TYPE "DT_PAR_GEN_MEAS_2"
VERSION : 0.1
   STRUCT
      OIL_NDE_TEMP_VAL_LOW { S7_SetPoint := 'False'} : "DT_PARAM_SOLO" := (FALSE, 320, 0, 0.0, 0, T#0MS, 0.0, 0.0, '°C');
      OIL_NDE_TEMP_VAL_HIGH { S7_SetPoint := 'False'} : "DT_PARAM_SOLO" := (FALSE, 321, 0, 150.0, 0, T#0MS, 0.0, 0.0, '°C');
      OIL_NDE_TEMP_SCAL_FACTOR { S7_SetPoint := 'False'} : "DT_PARAM_SOLO" := (FALSE, 322, 0, 1.0, 0, T#0MS, 0.0, 0.0, '°C');
      OIL_NDE_TEMP_OFFSET { S7_SetPoint := 'False'} : "DT_PARAM_SOLO" := (FALSE, 323, 0, 0.0, 0, T#0MS, 0.0, 0.0, '°C');
      OIL_NDE_TEMP_H { S7_SetPoint := 'False'} : "DT_PARAM_SOLO" := (FALSE, 324, 0, 120.0, 0, T#0MS, 0.0, 0.0, '°C');
      OIL_NDE_TEMP_HH { S7_SetPoint := 'False'} : "DT_PARAM_SOLO" := (FALSE, 325, 0, 130.0, 0, T#0MS, 0.0, 0.0, '°C');
      THRUST_NDE_TEMP_VAL_LOW { S7_SetPoint := 'False'} : "DT_PARAM_SOLO" := (FALSE, 326, 0, 1.0, 0, T#0MS, 0.0, 0.0, '°C');
      THRUST_NDE_TEMP_VAL_HIGH { S7_SetPoint := 'False'} : "DT_PARAM_SOLO" := (FALSE, 327, 0, 0.0, 0, T#0MS, 0.0, 0.0, '°C');
      THRUST_NDE_TEMP_SCAL_FACTOR { S7_SetPoint := 'False'} : "DT_PARAM_SOLO" := (FALSE, 328, 0, 1.0, 0, T#0MS, 0.0, 0.0, '°C');
      THRUST_NDE_TEMP_OFFSET { S7_SetPoint := 'False'} : "DT_PARAM_SOLO" := (FALSE, 329, 0, 0.0, 0, T#0MS, 0.0, 0.0, '°C');
      THRUST_NDE_TEMP_H { S7_SetPoint := 'False'} : "DT_PARAM_SOLO" := (FALSE, 330, 0, 70.0, 0, T#0MS, 0.0, 0.0, '°C');
      THRUST_NDE_TEMP_HH { S7_SetPoint := 'False'} : "DT_PARAM_SOLO" := (FALSE, 331, 0, 80.0, 0, T#0MS, 0.0, 0.0, '°C');
      PARAM_12 { S7_SetPoint := 'False'} : "DT_PARAM_SOLO" := (FALSE, 332, 0, 0.0, 0, T#0MS, 0.0, 0.0, '');
      PARAM_13 { S7_SetPoint := 'False'} : "DT_PARAM_SOLO" := (FALSE, 333, 0, 120.0, 0, T#0MS, 0.0, 0.0, '');
      PARAM_14 { S7_SetPoint := 'False'} : "DT_PARAM_SOLO" := (FALSE, 334, 0, 1.0, 0, T#0MS, 0.0, 0.0, '');
      PARAM_15 { S7_SetPoint := 'False'} : "DT_PARAM_SOLO" := (FALSE, 335, 0, 0.0, 0, T#0MS, 0.0, 0.0, '');
      PARAM_16 { S7_SetPoint := 'False'} : "DT_PARAM_SOLO" := (FALSE, 336, 0, 70.0, 0, T#0MS, 0.0, 0.0, '');
      PARAM_17 { S7_SetPoint := 'False'} : "DT_PARAM_SOLO" := (FALSE, 337, 0, 80.0, 0, T#0MS, 0.0, 0.0, '');
      PARAM_18 { S7_SetPoint := 'False'} : "DT_PARAM_SOLO" := (FALSE, 338, 0, 0.0, 0, T#0MS, 0.0, 0.0, '');
      PARAM_19 { S7_SetPoint := 'False'} : "DT_PARAM_SOLO" := (FALSE, 339, 0, 0.0, 0, T#0MS, 0.0, 0.0, '');
      PARAM_20 { S7_SetPoint := 'False'} : "DT_PARAM_SOLO" := (FALSE, 340, 0, 0.0, 0, T#0MS, 0.0, 0.0, '');
      PARAM_21 { S7_SetPoint := 'False'} : "DT_PARAM_SOLO" := (FALSE, 341, 0, 0.0, 0, T#0MS, 0.0, 0.0, '');
      PARAM_22 { S7_SetPoint := 'False'} : "DT_PARAM_SOLO" := (FALSE, 342, 0, 0.0, 0, T#0MS, 0.0, 0.0, '');
      PARAM_23 { S7_SetPoint := 'False'} : "DT_PARAM_SOLO" := (FALSE, 343, 0, 0.0, 0, T#0MS, 0.0, 0.0, '');
      PARAM_24 { S7_SetPoint := 'False'} : "DT_PARAM_SOLO" := (FALSE, 344, 0, 0.0, 0, T#0MS, 0.0, 0.0, '');
      PARAM_25 { S7_SetPoint := 'False'} : "DT_PARAM_SOLO" := (FALSE, 345, 0, 0.0, 0, T#0MS, 0.0, 0.0, '');
      PARAM_26 { S7_SetPoint := 'False'} : "DT_PARAM_SOLO" := (FALSE, 346, 0, 0.0, 0, T#0MS, 0.0, 0.0, '');
      PARAM_27 { S7_SetPoint := 'False'} : "DT_PARAM_SOLO" := (FALSE, 347, 0, 0.0, 0, T#0MS, 0.0, 0.0, '');
      PARAM_28 { S7_SetPoint := 'False'} : "DT_PARAM_SOLO" := (FALSE, 348, 0, 0.0, 0, T#0MS, 0.0, 0.0, '');
      PARAM_29 { S7_SetPoint := 'False'} : "DT_PARAM_SOLO" := (FALSE, 349, 0, 0.0, 0, T#0MS, 0.0, 0.0, '');
      PARAM_30 { S7_SetPoint := 'False'} : "DT_PARAM_SOLO" := (FALSE, 350, 0, 0.0, 0, T#0MS, 0.0, 0.0, '');
      PARAM_31 { S7_SetPoint := 'False'} : "DT_PARAM_SOLO" := (FALSE, 351, 0, 0.0, 0, T#0MS, 0.0, 0.0, '');
   END_STRUCT;

END_TYPE

